// TIA Portal project "Simatin1200_Coolmay_SCL" (V18)

(* hardware
DEVICE "S7-1200 station_1"  S7-1200 Station
   slot 0: "Rack_0"  S7-1200 Rack  Rack  V1.0
   slot 1: "PLC_1"  CPU 1215C DC/DC/Rly  6ES7 215-1HG40-0XB0  V4.5
   slot 101: "CM 1241 (RS422/485)_1"  6ES7 241-1CH32-0XB0  V2.2
*)

// ===== PLC "PLC_1"  CPU 1215C DC/DC/Rly =====

VAR_GLOBAL   // PLC tag table "Default tag table"
   "System_Byte" AT %MB1 : Byte;
   "FirstScan" AT %M1.0 : Bool;
   "DiagStatusUpdate" AT %M1.1 : Bool;
   "AlwaysTRUE" AT %M1.2 : Bool;
   "AlwaysFALSE" AT %M1.3 : Bool;
   "Clock_Byte" AT %MB0 : Byte;
   "Clock_10Hz" AT %M0.0 : Bool;
   "Clock_5Hz" AT %M0.1 : Bool;
   "Clock_2.5Hz" AT %M0.2 : Bool;
   "Clock_2Hz" AT %M0.3 : Bool;
   "Clock_1.25Hz" AT %M0.4 : Bool;
   "Clock_1Hz" AT %M0.5 : Bool;
   "Clock_0.625Hz" AT %M0.6 : Bool;
   "Clock_0.5Hz" AT %M0.7 : Bool;
   "Tag_MotorOnOff" AT %Q0.0 : Bool;
   "analogInput_1" AT %IW64 : Int;
   "analogInput_2" AT %IW66 : Int;
END_VAR

DATA_BLOCK "DB_HMI_Data"   // DB1
{ S7_Optimized_Access := 'TRUE' }
VERSION : 0.1
   VAR
      motorForwardOn : Bool;
      motorReversOn : Bool;
      motorStop : Bool;
      frequencySetpoint : Real;
      frequencyActual : Real;
      voltageOut : Real;
      currentOut : Real;
      MinValueClamp : Int;
      MaxValueClamp : Int;
      frequencySource : Int;
      sensorOn : Bool;
      timerDelayMotorSensorsOn : Time;
   END_VAR
BEGIN
END_DATA_BLOCK

DATA_BLOCK "DB_App"   // DB2
{ S7_Optimized_Access := 'TRUE' }
VERSION : 0.1
// stored: InstanceOfName FB_App
"FB_App"
BEGIN
END_DATA_BLOCK

DATA_BLOCK "TEST_OPC_UA"   // DB3
{ S7_Optimized_Access := 'TRUE' }
VERSION : 0.1
   VAR
      Static_1 : Real := 1.0;
      TEMP_1 : Real := 2.0;
      TEMP_2 : Real := 3.0;
      TEMP_3 : Real := 4.0;
      TEMP_4 : Real := 5.0;
      TEMP_5 : Real := 6.0;
      TEMP_6 : Real := 7.0;
   END_VAR
BEGIN
END_DATA_BLOCK

DATA_BLOCK "DB_MB_Comm_LoadConfig"   // DB5
{ S7_Optimized_Access := 'TRUE' }
VERSION : 0.1
   VAR
      BAUD : UDInt := 9600;
      PARITY : UInt;
      FLOW_CTRL : UInt;
      RTS_ON_DLY : UInt;
      RTS_OFF_DLY : UInt;
      RESP_TO : UInt := 1000;
      DONE : Bool;
      ERROR : Bool;
      STATUS : Word;
   END_VAR
BEGIN
END_DATA_BLOCK

DATA_BLOCK "DB_MB_TCP_ServerConfig"   // DB6
{ S7_Optimized_Access := 'FALSE' }
VERSION : 0.1
   VAR
      Connect : TCON_IP_v4;
      MB_Disconnect : Bool;
      MB_NDR : Bool;
      MB_DR : Bool;
      MB_Error : Bool;
      MB_Status : Word;
      HoldingReg : Array[0..20] of Word;
   END_VAR
BEGIN
   Connect.ConnectionType := 11;
   Connect.RemoteAddress.ADDR[1] := 0;
   Connect.RemoteAddress.ADDR[2] := 0;
   Connect.RemoteAddress.ADDR[3] := 0;
   Connect.RemoteAddress.ADDR[4] := 0;
   Connect.LocalPort := 502;
   Connect.InterfaceId := 64;
   Connect.ID := 1;
   // HoldingReg[0] : MotorOn_Cmd (0=Stop, <>0=Start)
   // HoldingReg[1] : SetFrequency_Hold
   // HoldingReg[2] : FrequencyAct_Hold
   // HoldingReg[3] : MinValueClamp
   // HoldingReg[4] : MaxValueClamp
   // HoldingReg[5] : frequencySource (Выбор источника задания частоты)
END_DATA_BLOCK

DATA_BLOCK "DB_VFD_Data"   // DB8
{ S7_Optimized_Access := 'FALSE' }
VERSION : 0.1
   VAR
      ReadRegs : Array[0..15] of Word;
      forward : Bool;
      revers : Bool;
      stop : Bool;
      setFrequency : Real;   // 0020h - 40033
      outputFrequency : Real;   // 0021h - 40034 actual
      outputCurrent : Real;   // 0022h - 40035
      outputVoltage : Real;   // 0025h - 40038
      voltageZPT : Int;   // 0026h - 40039
      statusInputTerminals : Int;   // 0029h - 40042
      commands : Int;   // 0000h - 40001
      settingFrequency : Int;   // 0001h - 40002
   END_VAR
BEGIN
END_DATA_BLOCK

DATA_BLOCK "DB_MB_RTU_MasterConfig"   // DB10
{ S7_Optimized_Access := 'TRUE' }
VERSION : 0.1
   VAR
      REQ : Bool;
      MB_ADDR : UInt := 1;
      MODE : USInt;
      DATA_ADDR : UDInt;
      DATA_LEN : UInt;
      DONE : Bool;
      BUSY : Bool;
      ERROR : Bool;
      STATUS : Word;
      ptrAddr : Int;
      "Step" : Int;
      StepRequest : Int;
   END_VAR
BEGIN
END_DATA_BLOCK

DATA_BLOCK "DB_Sensors"   // DB11
{ S7_Optimized_Access := 'TRUE' }
VERSION : 0.1
// stored: InstanceOfName FB_Sensors
"FB_Sensors"
BEGIN
END_DATA_BLOCK

FUNCTION_BLOCK "FB_App"   // FB1, SCL
{ S7_Optimized_Access := 'TRUE' }
VERSION : 0.1
   VAR
      frequencySource_Last : Int;
      frequencySetpoint_Last : Real;
      state_start : Bool := true;
      state_rev : Bool := true;
      state_stop : Bool := true;
   END_VAR
BEGIN

   "FC_ModbusSrv"();
   "FC_ModbusMaster"();
   "DB_Sensors"();


   // ПУСК РЕВЕРС СТОП. Можно добавить условие, если все флаги равны false, то поставить все флаги в true. Ну или хотя бы флаг стоп
   IF #state_start = false AND #state_rev = false AND #state_stop = false THEN
       #state_start := true;
       #state_rev := true;
       #state_stop := true;
   END_IF;
       IF "DB_MB_TCP_ServerConfig".HoldingReg[0].%X0 = 1 AND #state_start = TRUE THEN
       #state_start := false;
       "DB_MB_TCP_ServerConfig".HoldingReg[0].%X1 := false;
       "DB_MB_TCP_ServerConfig".HoldingReg[0].%X8 := false;
       "DB_MB_RTU_MasterConfig".StepRequest := 2;
       #state_rev := true;
       #state_stop := true;
       "DB_HMI_Data".motorForwardOn := true;
       "DB_HMI_Data".motorReversOn := false;
       "DB_HMI_Data".motorStop := false;
   END_IF;
   IF "DB_MB_TCP_ServerConfig".HoldingReg[0].%X1 = 1 AND #state_rev = TRUE THEN
       #state_rev := FALSE;
       "DB_MB_TCP_ServerConfig".HoldingReg[0].%X0 := false;
       "DB_MB_TCP_ServerConfig".HoldingReg[0].%X8 := false;
       "DB_MB_RTU_MasterConfig".StepRequest := 2;
       #state_start := TRUE;
       #state_stop := true;
       "DB_HMI_Data".motorForwardOn := FALSE;
       "DB_HMI_Data".motorReversOn := true;
       "DB_HMI_Data".motorStop := false;
   END_IF;
   IF "DB_MB_TCP_ServerConfig".HoldingReg[0].%X8 = 1 AND #state_stop = TRUE THEN
       #state_stop := false;
       "DB_MB_TCP_ServerConfig".HoldingReg[0].%X0 := false;
       "DB_MB_TCP_ServerConfig".HoldingReg[0].%X1 := false;
       "DB_MB_RTU_MasterConfig".StepRequest := 2;
       #state_start := TRUE;
       #state_rev := true;
       "DB_HMI_Data".motorForwardOn := false;
       "DB_HMI_Data".motorReversOn := false;
       "DB_HMI_Data".motorStop := true;
   END_IF;


   // УСТАВКА ЧАСТОТЫ
   // REAL -> два holding-регистра [1] и [2]
   "DB_HMI_Data".frequencySetpoint := DWORD_TO_REAL(SHL(IN := WORD_TO_DWORD("DB_MB_TCP_ServerConfig".HoldingReg[1]), N := 16) OR
                                                    WORD_TO_DWORD("DB_MB_TCP_ServerConfig".HoldingReg[2]));
   IF "DB_HMI_Data".frequencySetpoint <> #frequencySetpoint_Last THEN
       "DB_MB_RTU_MasterConfig".StepRequest := 3;
       #frequencySetpoint_Last := "DB_HMI_Data".frequencySetpoint;
   END_IF;

   // АКТУАЛЬНАЯ ЧАСТОТА
   // REAL -> два holding-регистра [3] и [4]
   "DB_MB_TCP_ServerConfig".HoldingReg[3] :=
   DWORD_TO_WORD(SHR(IN := REAL_TO_DWORD("DB_VFD_Data".outputFrequency), N:= 16));     // high word
   "DB_MB_TCP_ServerConfig".HoldingReg[4] :=
   DWORD_TO_WORD(REAL_TO_DWORD("DB_VFD_Data".outputFrequency) AND 16#FFFF);     // low word
   "DB_HMI_Data".frequencyActual := "DB_VFD_Data".outputFrequency;


   // ВЫБОР ИСТОЧНИКА ЗАДАНИЯ ЧАСТОТЫ
   // Int ->holding-регистр [5]
   "DB_HMI_Data".frequencySource := WORD_TO_INT("DB_MB_TCP_ServerConfig".HoldingReg[5]);
   IF "DB_HMI_Data".frequencySource <> #frequencySource_Last THEN
       "DB_MB_RTU_MasterConfig".StepRequest := 4;
       #frequencySource_Last := "DB_HMI_Data".frequencySource;
   END_IF;

   // ТОК
   // REAL -> Два holding-регистра [6] [7]
   "DB_MB_TCP_ServerConfig".HoldingReg[6] :=
   DWORD_TO_WORD(SHR(IN := REAL_TO_DWORD("DB_VFD_Data".outputCurrent), N:=16));
   "DB_MB_TCP_ServerConfig".HoldingReg[7] :=
   DWORD_TO_WORD(REAL_TO_DWORD("DB_VFD_Data".outputCurrent) AND 16#FFFF);
   "DB_HMI_Data".currentOut := "DB_VFD_Data".outputCurrent;

   // ВЫХОДНОЕ НАПРЯЖКНИЕ
   // Real -> Два holding-регистра [8] и [9]
   "DB_MB_TCP_ServerConfig".HoldingReg[8] :=
   DWORD_TO_WORD(SHR(IN := REAL_TO_DWORD("DB_VFD_Data".outputVoltage), N := 16));
   "DB_MB_TCP_ServerConfig".HoldingReg[9] :=
   DWORD_TO_WORD(REAL_TO_DWORD("DB_VFD_Data".outputVoltage) AND 16#FFFF);
   "DB_HMI_Data".voltageOut := "DB_VFD_Data".outputVoltage;

   // ВКЛ/ВЫКЛ ДАТЧИК holding-регистра [10] использую только 0 бит. Остальные в резерве 
   "DB_HMI_Data".sensorOn := "DB_MB_TCP_ServerConfig".HoldingReg[10].%X0;

   // ВРЕМЯ РАБОТЫ ДВИГАТЕЛЯ ПРИ СРАБАТЫВАНИИ ДАТЧИКА 
   //  holding-регистра [11] и [12]
   "DB_HMI_Data".timerDelayMotorSensorsOn := INT_TO_TIME(REAL_TO_INT((DWORD_TO_REAL(SHL(IN := WORD_TO_DWORD("DB_MB_TCP_ServerConfig".HoldingReg[11]), N := 16) OR
                                                           WORD_TO_DWORD("DB_MB_TCP_ServerConfig".HoldingReg[12])))*1000));
   "DB_Sensors".timeDelay := "DB_HMI_Data".timerDelayMotorSensorsOn;
END_FUNCTION_BLOCK

FUNCTION_BLOCK "FB_Sensors"   // FB2, SCL
{ S7_Optimized_Access := 'TRUE' }
VERSION : 0.1
   VAR
      voltage_HL : Real := 10.0;
      voltage_LL : Real := 0.0;
      distance_HL : Real := 1000.0;
      distance_LL : Real := 100.0;
      analogValue : Int;
      voltageOutput : Real;
      distanceOutput : Real;
      timeDelay : Time;
      "timer" : TP_TIME;
      trig : R_TRIG;
      startCond : Bool;
      state : Bool := true;
   END_VAR
BEGIN
   #analogValue := "analogInput_1";
   // напряжение 
   #voltageOutput := #analogValue * ((#voltage_HL - #voltage_LL) / 27648) + #voltage_LL;
   //Растояние 
   #distanceOutput := #analogValue * ((#distance_HL - #distance_LL) / 27648) + #distance_LL;



   IF "DB_HMI_Data".sensorOn THEN
       #startCond :=
       (#distanceOutput > 300.0) AND
       (#distanceOutput < 500.0) AND
       (NOT "DB_VFD_Data".forward) AND
       (NOT "DB_VFD_Data".revers);

       #trig(CLK := #startCond);
       #timer(
              IN := #trig.Q,
              PT := #timeDelay
       );
       IF #trig.Q AND #state THEN
           "DB_MB_TCP_ServerConfig".HoldingReg[0].%X0 := 1;
           "DB_MB_RTU_MasterConfig".StepRequest := 2;
           #state := false;
       END_IF;

       IF #timer.ET = #timer.PT AND NOT #state THEN
           "DB_MB_TCP_ServerConfig".HoldingReg[0].%X0 := 0;
           "DB_MB_TCP_ServerConfig".HoldingReg[0].%X8 := 1;
           "DB_MB_RTU_MasterConfig".StepRequest := 2;
           #state := true;
       END_IF;
   END_IF;
END_FUNCTION_BLOCK

FUNCTION "FC_ModbusMaster" : Void   // FC3, SCL
{ S7_Optimized_Access := 'TRUE' }
VERSION : 0.1
BEGIN

   // 1. Если блок свободен и нет активного запроса,
   //    выбираем шаг и сразу поднимаем REQ

   IF NOT "DB_MB_RTU_MasterConfig".BUSY
       AND NOT "DB_MB_RTU_MasterConfig".REQ THEN

       // Берём запрос из StepRequest
       "DB_MB_RTU_MasterConfig".Step := "DB_MB_RTU_MasterConfig".StepRequest;

       CASE "DB_MB_RTU_MasterConfig".Step OF

           0://чтение Регистров параметров монитора (0020h - 0029h)
               "DB_MB_RTU_MasterConfig".MODE := 0;
               "DB_MB_RTU_MasterConfig".DATA_ADDR := 40033;
               "DB_MB_RTU_MasterConfig".DATA_LEN := 10;
           1://чтение регистров команд (регистр 0000h и 0001h) 
               "DB_MB_RTU_MasterConfig".MODE := 0;
               "DB_MB_RTU_MasterConfig".DATA_ADDR := 40001;
               "DB_MB_RTU_MasterConfig".DATA_LEN := 2;
           2:// включение/выключение двигателя (запись в регистр 0000h значение 1)
               "DB_MB_RTU_MasterConfig".MODE := 1;
               "DB_MB_RTU_MasterConfig".DATA_ADDR := 40001;
               "DB_MB_RTU_MasterConfig".DATA_LEN := 1;
               "DB_VFD_Data".ReadRegs[0] := "DB_MB_TCP_ServerConfig".HoldingReg[0]; // MotorOn_Cmd (0=Stop, <>0=Start)

              // Измениеть предыдущую строку на присваивание значение из таблицы "DB_HMI_Data".MotorOn, А не из холдинг регистра

           3:// задание частоты (запись в регистр 0001h )
               "DB_MB_RTU_MasterConfig".MODE := 1;
               "DB_MB_RTU_MasterConfig".DATA_ADDR := 40002;
               "DB_MB_RTU_MasterConfig".DATA_LEN := 1;
               "DB_VFD_Data".ReadRegs[0] := INT_TO_WORD(REAL_TO_INT(("DB_HMI_Data".frequencySetpoint)*100));
           4:// выбор источника задания частоты (запись в регистр 2101h)
               "DB_MB_RTU_MasterConfig".MODE := 1;
               "DB_MB_RTU_MasterConfig".DATA_ADDR := 48450;
               "DB_MB_RTU_MasterConfig".DATA_LEN := 1;
               "DB_VFD_Data".ReadRegs[0] := "DB_MB_TCP_ServerConfig".HoldingReg[5];
           5:// (запись в регистр )
               "DB_MB_RTU_MasterConfig".MODE := 1;
               "DB_MB_RTU_MasterConfig".DATA_ADDR := 48450;
               "DB_MB_RTU_MasterConfig".DATA_LEN := 1;
               "DB_VFD_Data".ReadRegs[0] := "DB_MB_TCP_ServerConfig".HoldingReg[5];


           ELSE
               "DB_MB_RTU_MasterConfig".Step := 0;   // защита
       END_CASE;

       // Старт запроса
       "DB_MB_RTU_MasterConfig".REQ := TRUE;
   END_IF;

   // Завершение запроса (успешно)
   IF "DB_MB_RTU_MasterConfig".DONE THEN
       "DB_MB_RTU_MasterConfig".REQ := FALSE;

        // Запись значений регистров парамтров мониторинга в таблицу "DB_VFD_Data"
       CASE "DB_MB_RTU_MasterConfig".Step OF
           0:  // Считываем
               "DB_VFD_Data".setFrequency := (INT_TO_REAL(WORD_TO_INT("DB_VFD_Data".ReadRegs[0]))) / 100;
               "DB_VFD_Data".outputFrequency := (INT_TO_REAL(WORD_TO_INT("DB_VFD_Data".ReadRegs[1]))) / 100;
               "DB_VFD_Data".outputCurrent := (INT_TO_REAL(WORD_TO_INT("DB_VFD_Data".ReadRegs[2]))) / 10;
               "DB_VFD_Data".outputVoltage := (INT_TO_REAL(WORD_TO_INT("DB_VFD_Data".ReadRegs[5]))) / 10;
               "DB_VFD_Data".voltageZPT := WORD_TO_INT("DB_VFD_Data".ReadRegs[6]);
               "DB_VFD_Data".statusInputTerminals := WORD_TO_INT("DB_VFD_Data".ReadRegs[9]);


           1:  // читали 2 регистра другого типа
               "DB_VFD_Data".commands := WORD_TO_INT("DB_VFD_Data".ReadRegs[0]);
               "DB_VFD_Data".forward := "DB_VFD_Data".ReadRegs[0].%X0;
               "DB_VFD_Data".revers := "DB_VFD_Data".ReadRegs[0].%X1;
               IF "DB_VFD_Data".forward = false AND "DB_VFD_Data".revers = false THEN
                   "DB_VFD_Data".stop := true;
               ELSE
                   "DB_VFD_Data".stop := FALSE;
               END_IF;
               "DB_VFD_Data".settingFrequency := WORD_TO_INT("DB_VFD_Data".ReadRegs[1]);

       END_CASE;


       // case 1 -> 0 -> 1 -> 0 ->...
       IF "DB_MB_RTU_MasterConfig".Step >= 1 THEN
           IF "DB_MB_RTU_MasterConfig".Step = "DB_MB_RTU_MasterConfig".StepRequest THEN
               "DB_MB_RTU_MasterConfig".StepRequest := 0;
           END_IF;
       ELSE
           IF "DB_MB_RTU_MasterConfig".Step = "DB_MB_RTU_MasterConfig".StepRequest THEN
               "DB_MB_RTU_MasterConfig".StepRequest := "DB_MB_RTU_MasterConfig".Step + 1;
           END_IF;
       END_IF;


   END_IF;

   // Ошибка
   IF "DB_MB_RTU_MasterConfig".ERROR THEN
       "DB_MB_RTU_MasterConfig".REQ := FALSE;
       "DB_MB_RTU_MasterConfig".StepRequest := 0;   // на всякий случай
   END_IF;


   // формирование, отправка и прием запроса 
   "MB_MASTER_DB"(
                  REQ := "DB_MB_RTU_MasterConfig".REQ,
                  MB_ADDR := "DB_MB_RTU_MasterConfig".MB_ADDR,
                  MODE := "DB_MB_RTU_MasterConfig".MODE,
                  DATA_ADDR := "DB_MB_RTU_MasterConfig".DATA_ADDR,
                  DATA_LEN := "DB_MB_RTU_MasterConfig".DATA_LEN,
                  DONE => "DB_MB_RTU_MasterConfig".DONE,
                  BUSY => "DB_MB_RTU_MasterConfig".BUSY,
                  ERROR => "DB_MB_RTU_MasterConfig".ERROR,
                  STATUS => "DB_MB_RTU_MasterConfig".STATUS,
                  DATA_PTR := "DB_VFD_Data".ReadRegs
   );
END_FUNCTION

FUNCTION "FC_ModbusSrv" : Void   // FC4, SCL
{ S7_Optimized_Access := 'TRUE' }
VERSION : 0.1
BEGIN
   "MB_SERVER_DB"(DISCONNECT := "DB_MB_TCP_ServerConfig".MB_Disconnect,
                  NDR => "DB_MB_TCP_ServerConfig".MB_NDR,
                  DR => "DB_MB_TCP_ServerConfig".MB_DR,
                  ERROR => "DB_MB_TCP_ServerConfig".MB_Error,
                  STATUS => "DB_MB_TCP_ServerConfig".MB_Status,
                  MB_HOLD_REG := "DB_MB_TCP_ServerConfig".HoldingReg,
                  CONNECT := "DB_MB_TCP_ServerConfig".Connect);
END_FUNCTION

ORGANIZATION_BLOCK "Main"   // OB1, SCL, ProgramCycle
TITLE = "Main Program Sweep (Cycle)"
{ S7_Optimized_Access := 'TRUE' }
VERSION : 0.1
   VAR_INPUT
      Initial_Call : Bool;   // Initial call of this OB
      Remanence : Bool;   // =True, if remanent data are available
   END_VAR
BEGIN

   "MB_COMM_LOAD_DB"(
                     REQ:= NOT "DB_MB_Comm_LoadConfig".DONE AND NOT "DB_MB_Comm_LoadConfig".ERROR,
                     "PORT":="Local~CM_1241_(RS422_485)_1",
                     BAUD:="DB_MB_Comm_LoadConfig".BAUD,
                     PARITY:="DB_MB_Comm_LoadConfig".PARITY,
                     FLOW_CTRL:="DB_MB_Comm_LoadConfig".FLOW_CTRL,
                     RTS_ON_DLY:="DB_MB_Comm_LoadConfig".RTS_ON_DLY,
                     RTS_OFF_DLY:="DB_MB_Comm_LoadConfig".RTS_OFF_DLY,
                     RESP_TO:="DB_MB_Comm_LoadConfig".RESP_TO,
                     DONE=>"DB_MB_Comm_LoadConfig".DONE,
                     ERROR=>"DB_MB_Comm_LoadConfig".ERROR,
                     STATUS=>"DB_MB_Comm_LoadConfig".STATUS,
                     MB_DB:="MB_MASTER_DB");

   "DB_App"();
END_ORGANIZATION_BLOCK